Staubli VAL3: safeTemp.dtx

public sPoint sSPoint
  [0]
    bool bActive
    pointRx pPointRx
    string sName
public zoneItem zZoneItem
  [0]
    pointRx pO
    pointRx pX
    pointRx pY
    frame fBase
    pointRx pFirst
    pointRx pSecond
    bool bActive
    string sID
